// TIA Portal V20 export
// export: Created 2026-10-19T18:07:32.6342099Z, ExportSetting WithDefaults, DisplayName Totally Integrated Automation Portal, DisplayVersion V20 Update 6, DisplayName TIA Portal Openness, DisplayVersion V20 Update 6, DisplayName TIA Portal Version Control Interface, DisplayVersion V20 Update 6, DisplayName SINAMICS Startdrive Advanced, DisplayVersion V20 SP1, DisplayName SINAMICS Startdrive G130, G150, S120, S150, SINAMICS MV, G220, S200, S210, DisplayVersion V20 SP1, DisplayName SINAMICS Startdrive G110M, G120, G120C, G120D, G120P, G115D, DisplayVersion V20 SP1, DisplayName STEP 7 Professional, DisplayVersion V20 Update 6, DisplayName STEP 7 Safety, DisplayVersion V20 Update 2, DisplayName WinCC Basic/Comfort/Advanced, DisplayVersion V20 Update 6, DisplayName WinCC Unified, DisplayVersion V20 Update 6
DATA_BLOCK "SICK_Barcode_DB"   // DB47
VERSION : 0.1
// stored: AutoNumber true, DBAccessibleFromOPCUA true, DBAccessibleFromWebserver true, InstanceOfName SICK_Barcode_FB, InstanceOfType FB
"SICK_Barcode_FB"
   // VAR_INPUT
   //    Rd_Done : Bool;
   //    Req_Done : Bool;
   //    Req_Busy : Bool;
   //    Error : Bool;
   //    arrResult : Array[1..200] of Byte;
   //    iCounter : USInt;
   //    iLength : Int;
   //    Error_Code : DWord;
   // END_VAR
   // VAR_OUTPUT
   //    Test_Comm : Bool;
   //    Enable_Trigger : Bool;
   //    Disable_Trigger : Bool;
   //    Enable_Req : Bool;
   //    Result : String;
   //    Test_OK : Bool;
   // END_VAR
BEGIN
END_DATA_BLOCK
